(* IEC 61131-3 sources: PLC-Static-Analysis/modules/plc-rules/src/test/resources/PLCA-P001/locals, 1 file *)

(* ---- locals.st ---- *)
FUNCTION_BLOCK FB_L
VAR
    n : INT;
END_VAR
n := 1;
n := 2; // PLCA-P001
END_FUNCTION_BLOCK

FUNCTION F_L : INT
VAR
    n : INT;
END_VAR
n := 1;
n := 2;
F_L := n;
END_FUNCTION
